(* IEC 61131-3 sources: iolistgen/tests_support/pl_stub/src/DUTs/DigitalInput, 5 files *)

(* ---- E_DiAlarm.dut.st ---- *)
// Назначение: заглушка plc-process-lib 1.0.0 для проверки типов сгенерированного кода без CODESYS
//             (API.md, раздел 4.1); не библиотека — тел и внутренних переменных нет
// Автор:      kr0nsch
// Версия:     1.0.0 (выпуск библиотеки)
// Документ:   docs/GENERATORS.md, раздел «Проверка ST без CODESYS»
{attribute 'qualified_only'}
TYPE E_DiAlarm :
(
    State := 0,
    Failure := 1
) UINT;
END_TYPE

(* ---- E_DiFailValue.dut.st ---- *)
// Назначение: заглушка plc-process-lib 1.0.0 для проверки типов сгенерированного кода без CODESYS
//             (API.md, раздел 12.1); не библиотека — тел и внутренних переменных нет
// Автор:      kr0nsch
// Версия:     1.0.0 (выпуск библиотеки)
// Документ:   docs/GENERATORS.md, раздел «Проверка ST без CODESYS»
{attribute 'qualified_only'}
{attribute 'strict'}
TYPE E_DiFailValue :
(
    HoldLast := 0,
    ForceFalse := 1,
    ForceTrue := 2
) INT;
END_TYPE

(* ---- ST_DigitalInputCfg.dut.st ---- *)
// Назначение: заглушка plc-process-lib 1.0.0 для проверки типов сгенерированного кода без CODESYS
//             (API.md, раздел 12.1); не библиотека — тел и внутренних переменных нет
// Автор:      kr0nsch
// Версия:     1.0.0 (выпуск библиотеки)
// Документ:   docs/GENERATORS.md, раздел «Проверка ST без CODESYS»
{attribute 'qualified_only'}
TYPE ST_DigitalInputCfg :
STRUCT
    xInvert        : BOOL := FALSE;
    tOnDelay       : TIME := T#0S;
    tOffDelay      : TIME := T#0S;
    eFailValue     : E_DiFailValue := E_DiFailValue.HoldLast;
    xAlarmOnTrue   : BOOL := TRUE;
    tSubstMax      : TIME := T#8H;
    udiAlarmIdBase : UDINT := 0;
    // lint:allow STL007 имя массива по контракту API.md (префикс a + тип элемента)
    astAlarm       : ARRAY[0..GVL_Const.DEV_ALARMS_MAX - 1] OF ST_AlarmCfg := [
            (ePriority := E_AlarmPriority.None),
            (ePriority := E_AlarmPriority.Medium),
            (ePriority := E_AlarmPriority.None),
            (ePriority := E_AlarmPriority.None),
            (ePriority := E_AlarmPriority.None),
            (ePriority := E_AlarmPriority.None),
            (ePriority := E_AlarmPriority.None),
            (ePriority := E_AlarmPriority.None)];
END_STRUCT
END_TYPE

(* ---- ST_DigitalInputCmd.dut.st ---- *)
// Назначение: заглушка plc-process-lib 1.0.0 для проверки типов сгенерированного кода без CODESYS
//             (API.md, раздел 12.1); не библиотека — тел и внутренних переменных нет
// Автор:      kr0nsch
// Версия:     1.0.0 (выпуск библиотеки)
// Документ:   docs/GENERATORS.md, раздел «Проверка ST без CODESYS»
{attribute 'qualified_only'}
TYPE ST_DigitalInputCmd :
STRUCT
    stCommon    : ST_DeviceCmd;
    xSubstValue : BOOL;
END_STRUCT
END_TYPE

(* ---- ST_DigitalInputSts.dut.st ---- *)
// Назначение: заглушка plc-process-lib 1.0.0 для проверки типов сгенерированного кода без CODESYS
//             (API.md, раздел 12.1); не библиотека — тел и внутренних переменных нет
// Автор:      kr0nsch
// Версия:     1.0.0 (выпуск библиотеки)
// Документ:   docs/GENERATORS.md, раздел «Проверка ST без CODESYS»
{attribute 'qualified_only'}
TYPE ST_DigitalInputSts :
STRUCT
    stCommon        : ST_DeviceSts;
    uiSubstRemain_s : UINT;
END_STRUCT
END_TYPE
